// TIA Portal V20 export
Screen "Marriage_MB190_MB190R02"  1276x673
  ScreenItem "Rectangle_3" at 20,591 size 615x79  Type=HmiRectangle
  ScreenItem "Rectangle_5" at 648,67 size 605x40  Type=HmiRectangle
  ScreenItem "Casella di testo_26" at 23,6 size 1230x53  Type=HmiTextBox
  ScreenItem "Button_15" at 237,598 size 180x66  Type=HmiButton
  ScreenItem "Button_14" at 22,598 size 180x66  Type=HmiButton
  ScreenItem "Fusszeile_Button_ManualOPMode1_3" at 648,591 size 605x79  Type=HmiButton
  ScreenItem "Text_9" at 799,75 size 249x23  Type=HmiText
  ScreenItem "Rectangle_2" at 357,109 size 278x479  Type=HmiRectangle
  ScreenItem "Line_23" at 357,317 size 278x1  Type=HmiLine
  ScreenItem "Line_45" at 357,421 size 278x1  Type=HmiLine
  ScreenItem "Line_46" at 357,474 size 278x1  Type=HmiLine
  ScreenItem "Line_47" at 357,530 size 278x1  Type=HmiLine
  ScreenItem "Rectangle_6" at 357,67 size 278x40  Type=HmiRectangle
  ScreenItem "Text_10" at 398,75 size 195x28  Type=HmiText
  ScreenItem "Line_55" at 357,211 size 278x1  Type=HmiLine
  ScreenItem "Text_2" at 419,108 size 124x53  Type=HmiText
  ScreenItem "Circle_2" at 0,0 size 100x30  Type=HmiCircle
  ScreenItem "Circle_7" at 0,0 size 100x30  Type=HmiCircle
  ScreenItem "Text_15" at 419,158 size 158x53  Type=HmiText
  ScreenItem "Circle_8" at 0,0 size 100x30  Type=HmiCircle
  ScreenItem "Text_16" at 419,211 size 207x53  Type=HmiText
  ScreenItem "Circle_1" at 0,0 size 100x30  Type=HmiCircle
  ScreenItem "Text_1" at 419,264 size 124x53  Type=HmiText
  ScreenItem "Circle_9" at 0,0 size 100x30  Type=HmiCircle
  ScreenItem "Text_17" at 419,317 size 174x53  Type=HmiText
  ScreenItem "Circle_3" at 0,0 size 100x30  Type=HmiCircle
  ScreenItem "Text_3" at 419,369 size 124x53  Type=HmiText
  ScreenItem "Circle_4" at 0,0 size 100x30  Type=HmiCircle
  ScreenItem "Text_4" at 419,422 size 124x53  Type=HmiText
  ScreenItem "Circle_5" at 0,0 size 100x30  Type=HmiCircle
  ScreenItem "Text_5" at 419,474 size 124x53  Type=HmiText
  ScreenItem "Circle_6" at 0,0 size 100x30  Type=HmiCircle
  ScreenItem "Text_6" at 419,531 size 124x53  Type=HmiText
  ScreenItem "Line_1" at 358,369 size 278x1  Type=HmiLine
  ScreenItem "Line_2" at 352,264 size 278x1  Type=HmiLine
  ScreenItem "Line_3" at 360,159 size 278x1  Type=HmiLine
  ScreenItem "Rectangle_4" at 22,67 size 327x40  Type=HmiRectangle
  ScreenItem "Text_7" at 60,75 size 251x23  Type=HmiText
  ScreenItem "面板容器_1" at 131,107 size 220x219  Type=HmiFaceplateContainer
  ScreenItem "Button_26" at 22,110 size 108x23  Type=HmiButton
  ScreenItem "Button_7" at 22,134 size 108x21  Type=HmiButton
  ScreenItem "Button_2" at 22,154 size 108x21  Type=HmiButton
  ScreenItem "Button_1" at 22,175 size 108x21  Type=HmiButton
  ScreenItem "Button_4" at 22,194 size 108x21  Type=HmiButton
  ScreenItem "Button_6" at 22,234 size 108x21  Type=HmiButton
  ScreenItem "Button_8" at 22,256 size 108x21  Type=HmiButton
  ScreenItem "Button_9" at 22,277 size 108x21  Type=HmiButton
  ScreenItem "Button_24" at 22,215 size 108x21  Type=HmiButton
  ScreenItem "Button_31" at 22,299 size 108x21  Type=HmiButton
  ScreenItem "Rectangle_1" at 23,329 size 327x40  Type=HmiRectangle
  ScreenItem "Text_8" at 61,337 size 251x23  Type=HmiText
  ScreenItem "面板容器_2" at 131,370 size 220x219  Type=HmiFaceplateContainer
  ScreenItem "Button_3" at 23,372 size 108x23  Type=HmiButton
  ScreenItem "Button_5" at 23,396 size 108x21  Type=HmiButton
  ScreenItem "Button_10" at 23,416 size 108x21  Type=HmiButton
  ScreenItem "Button_11" at 23,437 size 108x21  Type=HmiButton
  ScreenItem "Button_12" at 23,456 size 108x21  Type=HmiButton
  ScreenItem "Button_13" at 23,496 size 108x21  Type=HmiButton
  ScreenItem "Button_16" at 23,518 size 108x21  Type=HmiButton
  ScreenItem "Button_17" at 23,539 size 108x21  Type=HmiButton
  ScreenItem "Button_18" at 23,477 size 108x21  Type=HmiButton
  ScreenItem "Button_19" at 23,561 size 108x21  Type=HmiButton
  ScreenItem "Title_OPOverview_ScreenOverview_X390_Y2_2" at 648,146 size 113x36  Type=HmiTextBox
  ScreenItem "Title_OPOverview_ScreenOverview_X390_Y2_4" at 772,146 size 111x36  Type=HmiTextBox
  ScreenItem "Title_OPOverview_ScreenOverview_X390_Y2_3" at 895,146 size 113x36  Type=HmiTextBox
  ScreenItem "Title_OPOverview_ScreenOverview_X390_Y2_1" at 1019,146 size 111x36  Type=HmiTextBox
  ScreenItem "Fusszeile_Button_ManualOPMode1_1" at 648,109 size 235x33  Type=HmiButton
  ScreenItem "Fusszeile_Button_ManualOPMode1_2" at 895,109 size 235x33  Type=HmiButton
  ScreenItem "IO field_1" at 648,187 size 113x36  Type=HmiIOField
  ScreenItem "Symbolic IO field_1" at 772,187 size 111x36  Type=HmiSymbolicIOField
  ScreenItem "IO field_20" at 895,187 size 113x36  Type=HmiIOField
  ScreenItem "Symbolic IO field_18" at 1019,187 size 111x36  Type=HmiSymbolicIOField
  ScreenItem "IO field_2" at 648,227 size 113x36  Type=HmiIOField
  ScreenItem "Symbolic IO field_2" at 772,227 size 111x36  Type=HmiSymbolicIOField
  ScreenItem "IO field_3" at 895,227 size 113x36  Type=HmiIOField
  ScreenItem "Symbolic IO field_3" at 1019,227 size 111x36  Type=HmiSymbolicIOField
  ScreenItem "IO field_4" at 648,268 size 113x36  Type=HmiIOField
  ScreenItem "Symbolic IO field_4" at 772,268 size 111x36  Type=HmiSymbolicIOField
  ScreenItem "IO field_5" at 895,268 size 113x36  Type=HmiIOField
  ScreenItem "Symbolic IO field_5" at 1019,268 size 111x36  Type=HmiSymbolicIOField
  ScreenItem "IO field_6" at 648,308 size 113x36  Type=HmiIOField
  ScreenItem "Symbolic IO field_6" at 772,308 size 111x36  Type=HmiSymbolicIOField
  ScreenItem "IO field_7" at 895,308 size 113x36  Type=HmiIOField
  ScreenItem "Symbolic IO field_7" at 1019,308 size 111x36  Type=HmiSymbolicIOField
  ScreenItem "IO field_8" at 648,349 size 113x36  Type=HmiIOField
  ScreenItem "Symbolic IO field_8" at 772,349 size 111x36  Type=HmiSymbolicIOField
  ScreenItem "IO field_9" at 895,349 size 113x36  Type=HmiIOField
  ScreenItem "Symbolic IO field_9" at 1019,349 size 111x36  Type=HmiSymbolicIOField
  ScreenItem "IO field_10" at 648,389 size 113x36  Type=HmiIOField
  ScreenItem "Symbolic IO field_10" at 772,389 size 111x36  Type=HmiSymbolicIOField
  ScreenItem "IO field_11" at 895,389 size 113x36  Type=HmiIOField
  ScreenItem "Symbolic IO field_11" at 1019,389 size 111x36  Type=HmiSymbolicIOField
  ScreenItem "IO field_12" at 648,430 size 113x36  Type=HmiIOField
  ScreenItem "Symbolic IO field_12" at 772,430 size 111x36  Type=HmiSymbolicIOField
  ScreenItem "IO field_13" at 895,430 size 113x36  Type=HmiIOField
  ScreenItem "Symbolic IO field_13" at 1019,430 size 111x36  Type=HmiSymbolicIOField
  ScreenItem "IO field_14" at 648,470 size 113x36  Type=HmiIOField
  ScreenItem "Symbolic IO field_14" at 772,470 size 111x36  Type=HmiSymbolicIOField
  ScreenItem "IO field_15" at 895,470 size 113x36  Type=HmiIOField
  ScreenItem "Symbolic IO field_15" at 1019,470 size 111x36  Type=HmiSymbolicIOField
  ScreenItem "IO field_16" at 648,511 size 113x36  Type=HmiIOField
  ScreenItem "Symbolic IO field_16" at 772,511 size 111x36  Type=HmiSymbolicIOField
  ScreenItem "IO field_17" at 895,511 size 113x36  Type=HmiIOField
  ScreenItem "Symbolic IO field_17" at 1019,511 size 111x36  Type=HmiSymbolicIOField
  ScreenItem "IO field_18" at 648,552 size 113x36  Type=HmiIOField
  ScreenItem "Symbolic IO field_19" at 772,552 size 111x36  Type=HmiSymbolicIOField
  ScreenItem "IO field_19" at 895,552 size 113x36  Type=HmiIOField
  ScreenItem "Symbolic IO field_20" at 1019,552 size 111x36  Type=HmiSymbolicIOField
  ScreenItem "Symbolic IO field_21" at 1142,187 size 111x36  Type=HmiSymbolicIOField
  ScreenItem "Symbolic IO field_22" at 1142,227 size 111x36  Type=HmiSymbolicIOField
  ScreenItem "Symbolic IO field_23" at 1142,268 size 111x36  Type=HmiSymbolicIOField
  ScreenItem "Symbolic IO field_24" at 1142,308 size 111x36  Type=HmiSymbolicIOField
  ScreenItem "Symbolic IO field_25" at 1142,349 size 111x36  Type=HmiSymbolicIOField
  ScreenItem "Symbolic IO field_26" at 1142,389 size 111x36  Type=HmiSymbolicIOField
  ScreenItem "Symbolic IO field_27" at 1142,430 size 111x36  Type=HmiSymbolicIOField
  ScreenItem "Symbolic IO field_28" at 1142,470 size 111x36  Type=HmiSymbolicIOField
  ScreenItem "Symbolic IO field_29" at 1142,511 size 111x36  Type=HmiSymbolicIOField
  ScreenItem "Symbolic IO field_30" at 1142,552 size 111x36  Type=HmiSymbolicIOField
  ScreenItem "Title_OPOverview_ScreenOverview_X390_Y2_5" at 1142,146 size 111x36  Type=HmiTextBox
  ScreenItem "Fusszeile_Button_ManualOPMode1_4" at 1142,109 size 111x33  Type=HmiButton
  ScreenItem "Button_20" at 453,598 size 180x66  Type=HmiButton
